Fanuc KAREL source: KB00034.KL

PROGRAM KB00034
%NOLOCKGROUP
%ENVIRONMENT STRNG
VAR
  P1: CONFIG
  P2: STRING[80]
BEGIN
  P2 = 'A'
  CNV_CONF_STR(P1, P2)
END KB00034
